RoboDK station: Pick and place(castillo).rdk

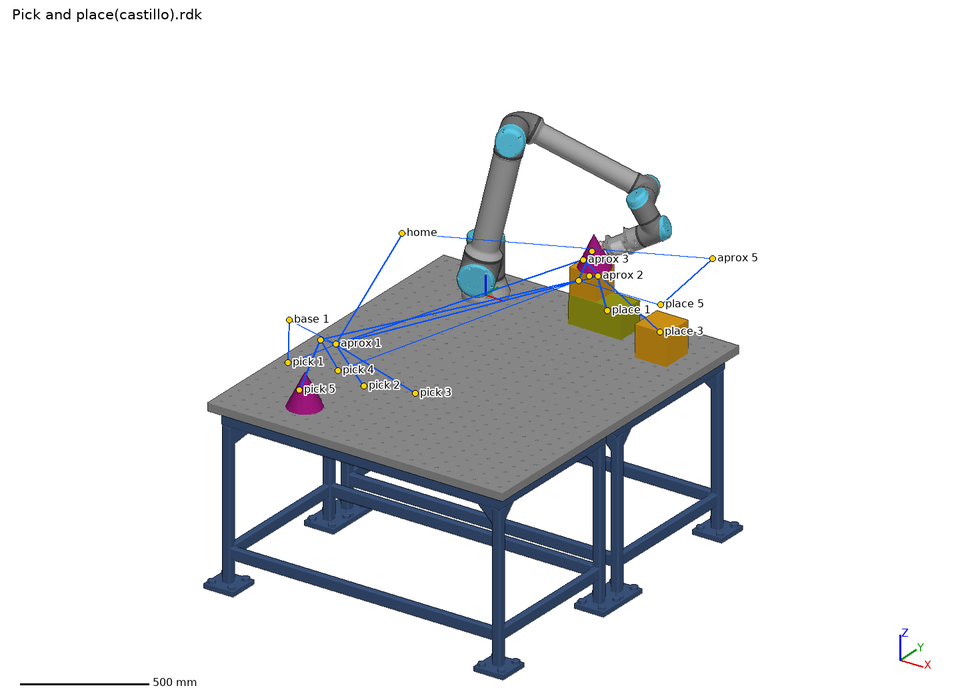
[picture v0: the station drawn from its stored meshes, robots at their saved joint values, targets as dots, program paths as lines]
Station Pick and place(castillo) (saved by RoboDK 6.1.1). Poses are relative to the parent item; angles as X-Y-Z fixed-axis rotations.
  - object Table 1400x800x800mm at (0, 800, 0) mm, size 1420 x 820 x 800 mm, geometry from Table-1400x800x800mm.sld
  - frame UR10e Base at (0, 1000, 0) mm
    - robot UR10e: 6 axes, payload 10 kg, reach 1300 mm, repeatability 0.05 mm, weight 28.9 kg
        modified DH rows (alpha deg, a mm, theta deg, d mm): 0, 0, 0, 180.7; 90, 0, 180, 0; 0, 612.6, 0, 0; 0, 571.335, 0, 174.15; -90, 0, 0, 119.85; 90, 0, 180, 116.55
        joint limits [-360, -360, -360, -360, -360, -360] to [360, 360, 360, 360, 360, 360]; home [0, -90, -90, 0, 90, 0]; saved at [25.894, -102.368, -104.43, -125.352, 94.636, 86.449]
      - tool SMC ZXP7A01-ZP25C-X1 Vacuum Gripper, TCP at (0, 0, 250) mm, size 88 x 106.8 x 127.9 mm
    - target home (Cartesian target) at (199.28, -848.63, 660.57) mm, rotated rx 178.13 ry -1.02 rz -139.96 deg; joints [-64.26, -112.93, -45.04, -113.59, 88.55, -14.26] of UR10e
    - target aprox 1  (Cartesian target) at (65.62, -1107.08, 249.11) mm, rotated rx -179.93 ry -1.51 rz -150.01 deg; joints [-76.734, -134.835, -52.261, -82.402, 88.571, -16.735] of UR10e
    - target base 1 (Cartesian target) at (-204.38, -1037.08, 249.11) mm, rotated rx -179.93 ry -1.51 rz -150.01 deg; joints [-90.467, -128.471, -63.289, -77.412, 88.731, -30.47] of UR10e
    - target pick 1 (Cartesian target) at (-204.38, -1047.08, 69.11) mm, rotated rx -179.93 ry -1.51 rz -150.01 deg; joints [-90.463, -135.316, -70.368, -63.489, 88.731, -30.466] of UR10e
    - target aprox 2 (Cartesian target) at (565.62, -47.08, 259.11) mm, rotated rx -179.93 ry -1.51 rz -150.01 deg; joints [10.632, -81.65, -121.899, -67.855, 89.433, 70.644] of UR10e
    - target place 1 (Cartesian target) at (546.58, 41.89, 68.32) mm, rotated rx -178.48 ry 0.07 rz 119.99 deg; joints [22.63, -89.676, -138.326, -43.496, 89.74, 172.647] of UR10e
    - target pick 2 (Cartesian target) at (155.62, -1047.08, 69.11) mm, rotated rx -179.93 ry -1.51 rz -150.01 deg; joints [-71.336, -135.189, -70.493, -63.951, 88.53, -11.335] of UR10e
    - target place 2 (Cartesian target) at (455.62, 52.92, 189.11) mm, rotated rx -179.93 ry -1.51 rz -150.01 deg; joints [25.092, -73.638, -135.68, -62.184, 89.801, 85.1] of UR10e
    - target pick 3 (Cartesian target) at (385.61, -1027.08, 95.11) mm, rotated rx -179.93 ry -1.51 rz -150.01 deg; joints [-59.877, -138.095, -62.225, -69.614, 88.487, 0.128] of UR10e
    - target aprox 3 (Cartesian target) at (565.62, -147.08, 369.11) mm, rotated rx -179.93 ry -1.51 rz -150.01 deg; joints [0.519, -81.249, -110.659, -79.375, 89.195, 60.534] of UR10e
    - target place 3 (Cartesian target) at (845.61, -27.08, 89.11) mm, rotated rx -179.93 ry -1.51 rz -150.01 deg; joints [8.343, -116.422, -100.201, -54.758, 89.377, 68.356] of UR10e
    - target aprox cone 1 (Cartesian target) at (48.71, -1186.61, 294.91) mm, rotated rx 145.9 ry -71.9 rz -123.09 deg; joints [-64.88, -141.6, -55.42, -86.5, 15.34, 3.62] of UR10e
    - target pick 4 (Cartesian target) at (-43.8, -934.63, 35.32) mm, rotated rx 168.01 ry -63.39 rz -146.05 deg; joints [-64.72, -132.153, -100.226, -47.151, 26.38, 4.67] of UR10e
    - target aprox cone 2 (Cartesian target) at (655.77, -307.37, 370.22) mm, rotated rx 168.77 ry -61.66 rz -146.63 deg; joints [-4.232, -120.003, -70.281, -139.602, 68.136, 71.815] of UR10e
    - target place 4 (Cartesian target) at (445.77, 82.63, 280.22) mm, rotated rx 168.77 ry -61.66 rz -146.63 deg; joints [25.894, -102.368, -104.43, -125.352, 94.636, 86.449] of UR10e
    - target pick 5 (Cartesian target) at (-45.58, -1195.93, 55.16) mm, rotated rx 152.47 ry -68.59 rz -129.01 deg; joints [-69.727, -152.201, -62.993, -50.51, 18.943, -14.815] of UR10e
    - target place 5 (Cartesian target) at (841.97, -16.57, 199.96) mm, rotated rx 151.45 ry -69.42 rz -125.54 deg; joints [12.75, -145.74, -46.93, -149, 79.03, 76.22] of UR10e
    - target aprox 5 (Cartesian target) at (1027.29, 69.15, 416.24) mm, rotated rx 179.98 ry 0.74 rz -152.15 deg; joints [11.9, -122.94, -55.41, -90.94, 90.22, 74.05] of UR10e
  - program armar castillo (45 instructions, listed below)
  - object Table 1400x800x800mm at (0, 0, 0) mm, size 1420 x 820 x 800 mm, geometry from Table-1400x800x800mm.sld
  - object Cone 500x500mm at (0, -200, 0) mm, size 149.2 x 150 x 150 mm, geometry from Cone-500x500mm.sld
  - object Prism 500x250x250mm at (533.1, 1034.98, -0.48) mm, rotated rx -0.47 ry -2.09 rz -89.98 deg, size 125 x 250 x 125 mm, geometry from Prism-500x250x250mm.sld
  - object Cube 50mm at (410, 980, 120) mm, size 125 x 125 x 125 mm, geometry from Cube-50mm.sld
  - object Cube 50mm at (790, 880, -6) mm, size 150 x 150 x 150 mm, geometry from Cube-50mm.sld
  - object Cone 500x500mm at (490.64, 1037.74, 245.64) mm, rotated rx 0.66 ry -1.63 rz 0.08 deg, size 139.3 x 140 x 140 mm, geometry from Cone-500x500mm.sld
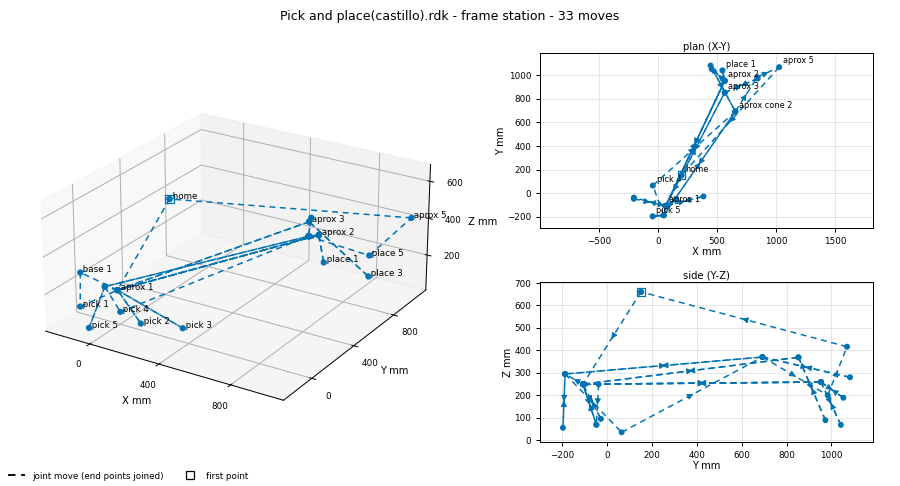
[picture p0: tool path of Pick and place(castillo).rdk in frame station, 33 of 33 moves have a stored position in this frame; points joined in program order, loops and branches not executed]

--- program armar castillo (robot UR10e) ---
  Est. Ref.: UR10e Base
  Mover objetos
  MoveJ (home)
  MoveJ (aprox 1 )
  MoveJ (base 1)
  MoveJ (pick 1)
  Adjuntar a SMC ZXP7A01-ZP25C-X1 Vacuum Gripper
  MoveJ (aprox 1 )
  MoveJ (aprox 2)
  MoveJ (place 1)
  Separar de SMC ZXP7A01-ZP25C-X1 Vacuum Gripper
  MoveJ (aprox 2)
  MoveJ (aprox 1 )
  MoveJ (pick 2)
  Adjuntar a SMC ZXP7A01-ZP25C-X1 Vacuum Gripper
  MoveJ (aprox 1 )
  MoveJ (aprox 2)
  MoveJ (place 2)
  Separar de SMC ZXP7A01-ZP25C-X1 Vacuum Gripper
  MoveJ (aprox 2)
  MoveJ (aprox 1 )
  MoveJ (pick 3)
  Adjuntar a SMC ZXP7A01-ZP25C-X1 Vacuum Gripper
  MoveJ (aprox 1 )
  MoveJ (aprox 3)
  MoveJ (place 3)
  Separar de SMC ZXP7A01-ZP25C-X1 Vacuum Gripper
  MoveJ (aprox 3)
  MoveJ (aprox 1 )
  MoveJ (aprox cone) -> target aprox cone 1
  MoveJ (pick 4)
  Adjuntar a SMC ZXP7A01-ZP25C-X1 Vacuum Gripper
  MoveJ (aprox cone) -> target aprox cone 2
  MoveJ (place 4)
  Separar de SMC ZXP7A01-ZP25C-X1 Vacuum Gripper
  MoveJ (aprox cone) -> target aprox cone 2
  MoveJ (aprox cone 1)
  MoveJ (pick 5)
  Adjuntar a SMC ZXP7A01-ZP25C-X1 Vacuum Gripper
  MoveJ (aprox cone 1)
  MoveJ (aprox cone 2)
  MoveJ (place 5)
  Separar de SMC ZXP7A01-ZP25C-X1 Vacuum Gripper
  MoveJ (aprox 5)
  MoveJ (home)
